// TwinCAT 3 PLC project CartonPLC
// ProgramVersion: 3.1.4026.28
// libraries:
//   SPT Base Types, 3.9.0 (Beckhoff Automation LLC)
//   Tc3_PackML_V2, * (Beckhoff Automation GmbH)
//   Tc3_EventLogger, * (Beckhoff Automation GmbH)
//   Tc2_System, * (Beckhoff Automation GmbH)
//   Tc3_Module, * (Beckhoff Automation GmbH)
//   Tc2_Standard, * (Beckhoff Automation GmbH)
// project tree:
//   / E_ConsoleCommand.TcDUT, GVL_HMI.TcGVL, FB_VirtualCylinder.TcPOU, FB_StrokeStation.TcPOU, FB_CartonCell.TcPOU, FB_SimAxis.TcPOU, FB_SealInspection.TcPOU, FB_CellDevices.TcPOU, I_LineClamp.TcIO, FB_LineClamp.TcPOU, FB_ContinuousLine.TcPOU, FB_LineEvents.TcPOU, MAIN.TcPOU, PlcTask.TcTTO
// real-time tasks:
//   TASK PlcTask: cycle T#10ms, priority 20, ADS port 350

CONFIGURATION CartonPLC
    RESOURCE PLC ON TwinCAT3
        TASK PlcTask(INTERVAL := T#10ms, PRIORITY := 20);
        PROGRAM MAIN WITH PlcTask : MAIN;
    END_RESOURCE
END_CONFIGURATION

// ---- E_ConsoleCommand.TcDUT
{attribute 'qualified_only'}
TYPE E_ConsoleCommand :
(
    Reset := 1,
    Start := 2,
    Hold := 3,
    Unhold := 4,
    Suspend := 5,
    Unsuspend := 6,
    Stop := 7,
    Abort := 8,
    Clear := 9,
    Automatic := 10,
    Manual := 11,
    Stroke1 := 12,
    Stroke2 := 13,
    Stroke3 := 14,
    Stroke4 := 15,
    Stroke5 := 16,
    DropAir := 17,
    RestoreAir := 18,
    LowBlanks := 19,
    Refill := 20,
    MissingSeal := 21,
    RestoreSeal := 22,
    LoopLine := 23,
    Bench := 24,
    Standard := 25,
    Precision := 26,
    JamClamp := 27,
    ReleaseClamp := 28,
    AckClamp := 29
) DINT;
END_TYPE

// ---- GVL_HMI.TcGVL
{attribute 'qualified_only'}
VAR_GLOBAL
    // One atomic DINT per request. See docs/ads.md for the word layout.
    Request : DINT;
    Status : ARRAY[0..105] OF DINT;
END_VAR

// ---- I_LineClamp.TcIO
INTERFACE I_LineClamp

METHOD Follow : DINT
VAR_INPUT
    Extend : BOOL;
END_VAR
END_METHOD

METHOD Home
END_METHOD

END_INTERFACE

// ---- MAIN.TcPOU
PROGRAM MAIN
VAR
    Cell : FB_CartonCell := (Name := 'Carton Cell');
END_VAR

Cell.RunScan();

END_PROGRAM

// ---- FB_CartonCell.TcPOU
FUNCTION_BLOCK FB_CartonCell EXTENDS SPT_BaseTypes.FB_PackML_BaseModule
VAR
    Line : FB_ContinuousLine;
    LineEvents : FB_LineEvents;
    Devices : FB_CellDevices;
    Stations : ARRAY[1..5] OF FB_StrokeStation;
    ActiveStation : DINT;
    Finished : BOOL;
    Cartons : DINT;
    AirFault : BOOL;
    LowStock : BOOL;
    PreviousState : Tc3_PackML_V2.E_PMLState;
    ActingScans : INT;
    RequestSample : DINT;
    Acknowledged : DINT;
    Accepted : BOOL;
    StatusBuffer : ARRAY[0..105] OF DINT;
END_VAR

METHOD PROTECTED Initialize : BOOL
// User mode 4 keeps Idle and Complete for one-station commissioning.
CustomModes(eMode := 4, sName := 'Manual stroke', bDisableHeld := TRUE,
    bDisableSuspended := TRUE, bEnableUnitModeChangeStopped := TRUE);
Initialize := SUPER^.Initialize();
END_METHOD

METHOD RunScan
IF _InitComplete THEN
    CyclicLogic();
ELSE
    _InitComplete := Initialize();
END_IF
END_METHOD

METHOD CyclicLogic
// SPT can call this hook while Initialize is still on the stack.
IF NOT _InitComplete THEN RETURN; END_IF

IF _CurrentState <> PreviousState THEN
    ActingScans := 0;
    PreviousState := _CurrentState;
ELSE
    ActingScans := MIN(45, ActingScans + 1);
END_IF

// Sample once so a concurrent ADS write belongs entirely to one scan.
RequestSample := GVL_HMI.Request;
IF RequestSample <> Acknowledged THEN
    Accepted := ApplyCommand(RequestSample MOD 256);
    Acknowledged := RequestSample;
END_IF

Line.Clock((_CurrentState = Tc3_PackML_V2.E_PMLState.ePMLState_Execute) AND Line.Enabled AND (_CurrentMode = E_PMLUnitMode.ePMLUnitMode_Production));
SUPER^.CyclicLogic();
LineEvents(Occurrence := Line.Occurrence, Alarm := Line.Alarm, Jammed := Line.Jammed,
    Idle := _CurrentState = Tc3_PackML_V2.E_PMLState.ePMLState_Idle);
PublishStatus();
END_METHOD

METHOD PROTECTED Execute
IF Line.Enabled AND (_CurrentMode = E_PMLUnitMode.ePMLUnitMode_Production) THEN
    IF Line.Alarm = 0 THEN Line.Step(Devices.MissingSeal); END_IF
    IF Line.Alarm <> 0 THEN ChangeState(Tc3_PackML_V2.E_PMLCommand.ePMLCommand_Abort); END_IF
    RETURN;
END_IF
IF (ActiveStation < 1) OR (ActiveStation > 5) THEN RETURN; END_IF
IF Finished THEN
    StateComplete();
    RETURN;
END_IF

Stations[ActiveStation].Step();
IF _CurrentMode = E_PMLUnitMode.ePMLUnitMode_Production THEN
    Devices.ProcessStation(ActiveStation, Stations[ActiveStation].Phase);
END_IF

IF Stations[ActiveStation].Done AND
   ((_CurrentMode = E_PMLUnitMode.ePMLUnitMode_UserMode1) OR Devices.ReadyToLeave(ActiveStation)) THEN
    IF (_CurrentMode = E_PMLUnitMode.ePMLUnitMode_UserMode1) OR (ActiveStation = 5) THEN
        Finished := TRUE;
        IF _CurrentMode = E_PMLUnitMode.ePMLUnitMode_Production THEN
            IF Devices.FinishCarton() THEN
                Cartons := Cartons + 1;
            END_IF
        END_IF
        StateComplete();
    ELSIF Devices.IndexToNext(ActiveStation) THEN
        ActiveStation := ActiveStation + 1;
    END_IF
END_IF
END_METHOD

METHOD PROTECTED Resetting
VAR
    StationIndex : INT;
END_VAR
FOR StationIndex := 1 TO 5 DO
    Stations[StationIndex].ResetStation();
END_FOR
Devices.ResetDevices();
Line.ResetLine();
ActiveStation := 0;
Finished := FALSE;
IF (_CurrentState = PreviousState) AND (ActingScans >= 45) THEN
    StateComplete();
END_IF
END_METHOD

METHOD PROTECTED Clearing
IF (_CurrentState = PreviousState) AND (ActingScans >= 45) THEN
    StateComplete();
END_IF
END_METHOD

METHOD PROTECTED Starting
IF (_CurrentState = PreviousState) AND (ActingScans >= 45) THEN
    StateComplete();
END_IF
END_METHOD

METHOD PROTECTED Stopping
IF (_CurrentState = PreviousState) AND (ActingScans >= 45) THEN
    StateComplete();
END_IF
END_METHOD

METHOD PROTECTED Aborting
IF (_CurrentState = PreviousState) AND (ActingScans >= 45) THEN
    StateComplete();
END_IF
END_METHOD

METHOD PROTECTED Holding
IF (_CurrentState = PreviousState) AND (ActingScans >= 45) THEN
    StateComplete();
END_IF
END_METHOD

METHOD PROTECTED Unholding
IF (_CurrentState = PreviousState) AND (ActingScans >= 45) THEN
    StateComplete();
END_IF
END_METHOD

METHOD PROTECTED Suspending
IF (_CurrentState = PreviousState) AND (ActingScans >= 45) THEN
    StateComplete();
END_IF
END_METHOD

METHOD PROTECTED Unsuspending
IF (_CurrentState = PreviousState) AND (ActingScans >= 45) THEN
    StateComplete();
END_IF
END_METHOD

METHOD PROTECTED Completing
IF (_CurrentState = PreviousState) AND (ActingScans >= 45) THEN
    StateComplete();
END_IF
END_METHOD

METHOD PRIVATE ApplyCommand : BOOL
VAR_INPUT
    Code : DINT;
END_VAR
VAR
    IsManual : BOOL;
END_VAR
IsManual := _CurrentMode = E_PMLUnitMode.ePMLUnitMode_UserMode1;
CASE Code OF
    E_ConsoleCommand.Reset:
        IF NOT AirFault AND ((_CurrentState = Tc3_PackML_V2.E_PMLState.ePMLState_Stopped) OR (_CurrentState = Tc3_PackML_V2.E_PMLState.ePMLState_Complete)) THEN
            ChangeState(Tc3_PackML_V2.E_PMLCommand.ePMLCommand_Reset);
            ApplyCommand := TRUE;
        END_IF
    E_ConsoleCommand.Start:
        IF NOT IsManual AND (_CurrentState = Tc3_PackML_V2.E_PMLState.ePMLState_Idle) THEN
            Line.Timing := Line.Enabled;
            ActiveStation := SEL(Line.Enabled, 1, 0);
            ChangeState(Tc3_PackML_V2.E_PMLCommand.ePMLCommand_Start);
            ApplyCommand := TRUE;
        END_IF
    E_ConsoleCommand.Hold:
        IF NOT IsManual AND (_CurrentState = Tc3_PackML_V2.E_PMLState.ePMLState_Execute) THEN
            ChangeState(Tc3_PackML_V2.E_PMLCommand.ePMLCommand_Hold);
            ApplyCommand := TRUE;
        END_IF
    E_ConsoleCommand.Unhold:
        IF _CurrentState = Tc3_PackML_V2.E_PMLState.ePMLState_Held THEN
            ChangeState(Tc3_PackML_V2.E_PMLCommand.ePMLCommand_Unhold);
            ApplyCommand := TRUE;
        END_IF
    E_ConsoleCommand.Suspend:
        IF NOT IsManual AND (_CurrentState = Tc3_PackML_V2.E_PMLState.ePMLState_Execute) THEN
            ChangeState(Tc3_PackML_V2.E_PMLCommand.ePMLCommand_Suspend);
            ApplyCommand := TRUE;
        END_IF
    E_ConsoleCommand.Unsuspend:
        IF _CurrentState = Tc3_PackML_V2.E_PMLState.ePMLState_Suspended THEN
            ChangeState(Tc3_PackML_V2.E_PMLCommand.ePMLCommand_Unsuspend);
            ApplyCommand := TRUE;
        END_IF
    E_ConsoleCommand.Stop:
        IF (_CurrentState <> Tc3_PackML_V2.E_PMLState.ePMLState_Undefined) AND
            (_CurrentState <> Tc3_PackML_V2.E_PMLState.ePMLState_Stopped) AND
            (_CurrentState <> Tc3_PackML_V2.E_PMLState.ePMLState_Stopping) AND
            (_CurrentState <> Tc3_PackML_V2.E_PMLState.ePMLState_Aborted) AND
            (_CurrentState <> Tc3_PackML_V2.E_PMLState.ePMLState_Aborting) AND
            (_CurrentState <> Tc3_PackML_V2.E_PMLState.ePMLState_Clearing) THEN
            Line.Timing := FALSE;
            ChangeState(Tc3_PackML_V2.E_PMLCommand.ePMLCommand_Stop);
            ApplyCommand := TRUE;
        END_IF
    E_ConsoleCommand.Abort:
        IF (_CurrentState <> Tc3_PackML_V2.E_PMLState.ePMLState_Aborted) AND
            (_CurrentState <> Tc3_PackML_V2.E_PMLState.ePMLState_Aborting) AND
            (_CurrentState <> Tc3_PackML_V2.E_PMLState.ePMLState_Undefined) THEN
            ChangeState(Tc3_PackML_V2.E_PMLCommand.ePMLCommand_Abort);
            ApplyCommand := TRUE;
        END_IF
    E_ConsoleCommand.Clear:
        IF NOT AirFault AND ((Line.Alarm = 0) OR ((Line.Alarm = 2) AND NOT Line.Jammed)) AND (_CurrentState = Tc3_PackML_V2.E_PMLState.ePMLState_Aborted) THEN
            Line.ClearAlarm();
            ChangeState(Tc3_PackML_V2.E_PMLCommand.ePMLCommand_Clear);
            ApplyCommand := TRUE;
        END_IF
    E_ConsoleCommand.Manual, E_ConsoleCommand.Automatic:
        IF _CurrentState = Tc3_PackML_V2.E_PMLState.ePMLState_Stopped THEN
            IF (Code = E_ConsoleCommand.Manual) AND NOT IsManual THEN
                Line.Timing := FALSE;
                ChangeMode(E_PMLUnitMode.ePMLUnitMode_UserMode1);
                ApplyCommand := TRUE;
            ELSIF (Code = E_ConsoleCommand.Automatic) AND IsManual THEN
                ChangeMode(E_PMLUnitMode.ePMLUnitMode_Production);
                ApplyCommand := TRUE;
            END_IF
        END_IF
    E_ConsoleCommand.Stroke1..E_ConsoleCommand.Stroke5:
        IF IsManual AND (_CurrentState = Tc3_PackML_V2.E_PMLState.ePMLState_Idle) THEN
            ActiveStation := Code - E_ConsoleCommand.Stroke1 + 1;
            ChangeState(Tc3_PackML_V2.E_PMLCommand.ePMLCommand_Start);
            ApplyCommand := TRUE;
        END_IF
    E_ConsoleCommand.DropAir:
        ApplyCommand := NOT AirFault;
        AirFault := TRUE;
        IF (_CurrentState <> Tc3_PackML_V2.E_PMLState.ePMLState_Aborted) AND (_CurrentState <> Tc3_PackML_V2.E_PMLState.ePMLState_Aborting) THEN
            ChangeState(Tc3_PackML_V2.E_PMLCommand.ePMLCommand_Abort);
        END_IF
    E_ConsoleCommand.RestoreAir:
        ApplyCommand := AirFault;
        AirFault := FALSE;
    E_ConsoleCommand.LowBlanks:
        ApplyCommand := NOT LowStock;
        LowStock := TRUE;
    E_ConsoleCommand.MissingSeal:
        ApplyCommand := NOT Devices.MissingSeal;
        Devices.MissingSeal := TRUE;
    E_ConsoleCommand.RestoreSeal:
        ApplyCommand := Devices.MissingSeal;
        Devices.MissingSeal := FALSE;
    E_ConsoleCommand.LoopLine, E_ConsoleCommand.Bench:
        IF NOT IsManual AND (_CurrentState = Tc3_PackML_V2.E_PMLState.ePMLState_Stopped) THEN
            ApplyCommand := Line.Enabled <> (Code = E_ConsoleCommand.LoopLine);
            Line.Timing := FALSE;
            Line.Enabled := Code = E_ConsoleCommand.LoopLine;
        END_IF
    E_ConsoleCommand.Standard, E_ConsoleCommand.Precision:
        IF Line.Enabled AND NOT IsManual AND (_CurrentState = Tc3_PackML_V2.E_PMLState.ePMLState_Stopped) THEN
            ApplyCommand := Line.Precision <> (Code = E_ConsoleCommand.Precision);
            Line.Precision := Code = E_ConsoleCommand.Precision;
        END_IF
    E_ConsoleCommand.JamClamp:
        IF Line.Enabled AND NOT IsManual AND NOT Line.Jammed AND (Line.Alarm = 0) THEN
            Line.Jammed := TRUE; ApplyCommand := TRUE;
        END_IF
    E_ConsoleCommand.ReleaseClamp:
        ApplyCommand := Line.Jammed; Line.Jammed := FALSE;
    E_ConsoleCommand.AckClamp:
        IF (_CurrentState = Tc3_PackML_V2.E_PMLState.ePMLState_Aborted) AND
            (Line.Alarm = 1) AND (RequestSample / 256 = Line.Occurrence) THEN
            Line.AcknowledgeAlarm(); ApplyCommand := TRUE;
        END_IF
    E_ConsoleCommand.Refill:
        ApplyCommand := LowStock;
        LowStock := FALSE;
END_CASE
END_METHOD

METHOD PRIVATE PublishStatus
StatusBuffer[0] := 51003;
StatusBuffer[1] := TO_DINT(_CurrentState);
StatusBuffer[2] := BOOL_TO_DINT(_CurrentMode = E_PMLUnitMode.ePMLUnitMode_UserMode1);
StatusBuffer[3] := ActiveStation;
StatusBuffer[4] := 0;
IF (ActiveStation >= 1) AND (ActiveStation <= 5) THEN
    StatusBuffer[4] := Stations[ActiveStation].Phase;
END_IF
StatusBuffer[5] := Cartons;
StatusBuffer[6] := BOOL_TO_DINT(AirFault);
StatusBuffer[7] := BOOL_TO_DINT(LowStock);
StatusBuffer[8] := Acknowledged;
StatusBuffer[9] := (StatusBuffer[9] MOD 2000000000) + 1;
StatusBuffer[10] := BOOL_TO_DINT(Accepted);
Devices.Publish(StatusBuffer);
Line.Publish(StatusBuffer);
GVL_HMI.Status := StatusBuffer;
END_METHOD

END_FUNCTION_BLOCK

// ---- FB_ContinuousLine.TcPOU
FUNCTION_BLOCK FB_ContinuousLine
VAR
    Clamp : FB_LineClamp;
    Actuator : I_LineClamp;
    Vision : FB_SealInspection;
    Products, Checks, Failures : ARRAY[0..15] OF DINT;
    CamX, CamZ : ARRAY[0..7] OF DINT;
    Tick, PitchIndex, Issued, Good, Rejected, LastId, LastFailed, LastChecked, Discarded : DINT;
    RunTicks, PlannedTicks, IdealTicks, WaitTicks, Travel, ClampMm : DINT;
    ClampRequest : BOOL;
END_VAR
VAR_INPUT
    Enabled : BOOL := TRUE;
    Precision, Jammed, Timing : BOOL;
END_VAR
VAR_OUTPUT
    Alarm, Occurrence : DINT;
END_VAR

METHOD ClearAlarm
Alarm := 0;
END_METHOD

METHOD AcknowledgeAlarm
Alarm := 2;
END_METHOD

METHOD Clock
VAR_INPUT
    Executing : BOOL;
END_VAR
IF Timing THEN
    PlannedTicks := PlannedTicks + 1;
    IF Executing THEN RunTicks := RunTicks + 1; END_IF
END_IF
END_METHOD

METHOD ResetLine
VAR
    i : INT;
END_VAR
FOR i := 0 TO 15 DO
    IF Products[i] <> 0 THEN Discarded := Discarded + 1; END_IF
    Products[i] := 0; Checks[i] := 0; Failures[i] := 0;
END_FOR
FOR i := 0 TO 7 DO CamX[i] := 0; CamZ[i] := 0; END_FOR
Tick := 0; PitchIndex := 0; WaitTicks := 0; Travel := 0;
Actuator := Clamp;
Actuator.Home();
ClampMm := 0; ClampRequest := FALSE;
END_METHOD

METHOD AtSlot : DINT
VAR_INPUT
    Slot, Count : DINT;
END_VAR
AtSlot := (Slot + Count - (PitchIndex MOD Count)) MOD Count;
END_METHOD

METHOD Ease : DINT
VAR_INPUT
    InputPhase : DINT;
END_VAR
VAR
    u : DINT;
END_VAR
u := LIMIT(0, InputPhase, 100);
Ease := u * u * (300 - 2 * u) / 1000;
END_METHOD

METHOD InspectMover
VAR_INPUT
    Mover, BitNumber : DINT;
    Passed : BOOL;
END_VAR
VAR
    Mask : DWORD;
END_VAR
Mask := SHL(DWORD#1, DINT_TO_UINT(BitNumber));
Checks[Mover] := DWORD_TO_DINT(DINT_TO_DWORD(Checks[Mover]) OR Mask);
IF NOT Passed THEN Failures[Mover] := DWORD_TO_DINT(DINT_TO_DWORD(Failures[Mover]) OR Mask); END_IF
END_METHOD

METHOD Step
VAR_INPUT
    MissingSeal : BOOL;
END_VAR
VAR
    p, Mover, Station, Reach, Depth, Stroke : DINT;
    FirstScan : BOOL;
END_VAR
VAR CONSTANT
    Period : DINT := 200; // 2 s at the 10 ms scan rate
END_VAR
Stroke := SEL(Precision, 40, 48);
p := Tick * 100 / Period;
FirstScan := (Tick MOD (Period / 100)) = 0;
Mover := AtSlot(0, 10);
IF (Tick = 0) AND (Products[Mover] = 0) THEN
    Issued := Issued + 1; Products[Mover] := Issued;
END_IF
ClampRequest := (Products[AtSlot(2, 10)] <> 0) AND (p >= 12) AND (p < 54);
Actuator := Clamp;
Clamp.Jammed := Jammed;
ClampMm := Actuator.Follow(ClampRequest);
IF ClampRequest AND (ClampMm < 16) THEN WaitTicks := WaitTicks + 1; ELSE WaitTicks := 0; END_IF
IF WaitTicks >= 15 THEN
    Occurrence := (Occurrence MOD 8388606) + 1;
    Alarm := 1;
    RETURN;
END_IF
IF p < 12 THEN Reach := Ease(p * 100 / 12);
ELSIF p < 48 THEN Reach := 1000;
ELSE Reach := 1000 - Ease((p - 48) * 100 / 12); END_IF
IF p < 12 THEN Depth := 0;
ELSIF p < 26 THEN Depth := Ease((p - 12) * 100 / 14);
ELSIF p < 36 THEN Depth := 1000;
ELSE Depth := 1000 - Ease((p - 36) * 100 / 12); END_IF
Travel := Ease((p - 60) * 100 / 40);
FOR Station := 0 TO 7 DO
    Mover := AtSlot(SEL(Station < 4, Station + 1, Station), 10);
    IF Products[Mover] <> 0 THEN
        CamX[Station] := Reach * (100 + Station * 4) / 1000;
        CamZ[Station] := Depth * Stroke / 1000;
        IF Station = 5 THEN
            IF p <= 80 THEN CamX[Station] := Travel / 2;
            ELSE CamX[Station] := 250 - Ease((p-80)*100/20) / 4; END_IF
            IF p < 60 THEN CamZ[Station] := 0;
            ELSIF p <= 74 THEN CamZ[Station] := Ease((p-60)*100/14) * Stroke / 1000;
            ELSE CamZ[Station] := (1000-Ease((p-78)*100/8)) * Stroke / 1000; END_IF
        END_IF
        IF (p = SEL(Station = 5, 32, 76)) AND FirstScan THEN
            InspectMover(Mover, Station, (CamZ[Station] = Stroke) AND ((Station <> 2) OR (ClampMm = 16)));
        END_IF
    ELSE CamX[Station] := 0; CamZ[Station] := 0; END_IF
END_FOR
IF (p = 54) AND FirstScan THEN ProcessTable(MissingSeal, Period); END_IF
Tick := Tick + 1;
IF Tick = Period THEN
    Tick := 0; Travel := 0; PitchIndex := (PitchIndex + 1) MOD 30;
END_IF
END_METHOD

METHOD ProcessTable
VAR_INPUT
    MissingSeal : BOOL;
    Period : DINT;
END_VAR
VAR
    Source, Target, Seat, Camera, Pack : DINT;
END_VAR
Source := AtSlot(8,10); Target := 10 + AtSlot(0,6);
IF (Products[Source] <> 0) AND (Products[Target] = 0) THEN
    Products[Target] := Products[Source]; Checks[Target] := Checks[Source]; Failures[Target] := Failures[Source];
    Products[Source] := 0; Checks[Source] := 0; Failures[Source] := 0;
END_IF
Seat := 10 + AtSlot(1,6); Camera := 10 + AtSlot(2,6); Pack := 10 + AtSlot(3,6);
IF Products[Seat] <> 0 THEN InspectMover(Seat, 8, (DINT_TO_DWORD(Checks[Seat]) AND DWORD#255) = DWORD#255); END_IF
IF Products[Camera] <> 0 THEN
    Vision.ClearResult(); Vision.Inspect(MissingSeal);
    InspectMover(Camera, 9, Vision.Verdict = 1);
END_IF
IF Products[Pack] <> 0 THEN
    LastId := Products[Pack]; LastChecked := Checks[Pack]; LastFailed := Failures[Pack];
    IF (LastChecked = 1023) AND (LastFailed = 0) THEN Good := Good + 1;
    ELSE Rejected := Rejected + 1; END_IF
    IdealTicks := IdealTicks + Period;
    Products[Pack] := 0; Checks[Pack] := 0; Failures[Pack] := 0;
END_IF
END_METHOD

METHOD Publish
VAR_IN_OUT
    Words : ARRAY[0..105] OF DINT;
END_VAR
VAR
    i : INT;
END_VAR
Words[20] := BOOL_TO_DINT(Enabled);
Words[21] := BOOL_TO_DINT(Precision);
Words[22] := Tick;
Words[23] := PitchIndex;
Words[24] := Issued;
Words[25] := Good;
Words[26] := Rejected;
Words[27] := LastId;
Words[28] := LastFailed;
Words[29] := BOOL_TO_DINT(Jammed);
Words[30] := Occurrence;
Words[31] := Alarm;
Words[32] := BOOL_TO_DINT(ClampRequest);
Words[33] := ClampMm;
Words[34] := RunTicks;
Words[35] := PlannedTicks;
Words[36] := IdealTicks;
Words[37] := Discarded;
FOR i := 0 TO 15 DO
    Words[40+i] := Products[i]; Words[56+i] := Checks[i]; Words[72+i] := Failures[i];
END_FOR
FOR i := 0 TO 7 DO Words[88+i] := CamX[i]; Words[96+i] := CamZ[i]; END_FOR
Words[104] := Travel;
Words[105] := LastChecked;
END_METHOD

END_FUNCTION_BLOCK

// ---- FB_LineClamp.TcPOU
FUNCTION_BLOCK FB_LineClamp IMPLEMENTS I_LineClamp
VAR_INPUT
    Jammed : BOOL;
END_VAR
VAR
    Position : DINT;
END_VAR

METHOD Follow : DINT
VAR_INPUT
    Extend : BOOL;
END_VAR
IF NOT Extend THEN Position := MAX(0, Position - 4);
ELSIF NOT Jammed THEN Position := MIN(16, Position + 4);
END_IF
Follow := Position;
END_METHOD

METHOD Home
Position := 0;
END_METHOD

END_FUNCTION_BLOCK

// ---- FB_SealInspection.TcPOU
FUNCTION_BLOCK FB_SealInspection
VAR_OUTPUT
    Verdict : DINT; // 0 pending, 1 pass, 2 reject
    BrightSamples : DINT;
END_VAR
VAR CONSTANT
    GoodPixels : ARRAY[0..4] OF USINT := [231, 236, 228, 239, 232];
    MissingPixels : ARRAY[0..4] OF USINT := [118, 122, 120, 124, 121];
END_VAR

METHOD Inspect
VAR_INPUT
    MissingSeal : BOOL;
END_VAR
VAR
    Index : INT;
    Pixel : USINT;
END_VAR
IF Verdict <> 0 THEN RETURN; END_IF
FOR Index := 0 TO 4 DO
    Pixel := SEL(MissingSeal, GoodPixels[Index], MissingPixels[Index]);
    IF Pixel >= 200 THEN
        BrightSamples := BrightSamples + 1;
    END_IF
END_FOR
Verdict := SEL(BrightSamples >= 4, 2, 1);
END_METHOD

METHOD ClearResult
Verdict := 0;
BrightSamples := 0;
END_METHOD

END_FUNCTION_BLOCK

// ---- FB_LineEvents.TcPOU
FUNCTION_BLOCK FB_LineEvents
VAR_INPUT
    Occurrence, Alarm : DINT;
    Jammed, Idle : BOOL;
END_VAR
VAR
    Event : Tc3_EventLogger.FB_TcAlarm;
    Recovery : Tc3_EventLogger.FB_TcMessage;
    Created, MessageCreated, Confirmed, Cleared, Recovered : BOOL;
    Seen : DINT;
END_VAR

IF NOT Created THEN Created := Event.CreateEx(TC_EVENTS.CartonLine.ClampTimeout, TRUE, 0) = 0; END_IF
IF NOT MessageCreated THEN MessageCreated := Recovery.CreateEx(TC_EVENTS.CartonLine.LineRecovered, 0) = 0; END_IF
IF Created AND (Occurrence <> Seen) THEN
    Event.ipArguments.Clear().AddDInt(Occurrence);
    IF Event.Raise(0) = 0 THEN Seen := Occurrence; Confirmed := FALSE; Cleared := FALSE; Recovered := FALSE; END_IF
END_IF
IF (Seen <> 0) AND (Seen = Occurrence) THEN
    IF (Alarm = 2) AND NOT Confirmed THEN Confirmed := Event.Confirm(0) = 0; END_IF
    IF NOT Jammed AND NOT Cleared THEN Cleared := Event.Clear(0, FALSE) = 0; END_IF
    IF MessageCreated AND Idle AND (Alarm = 0) AND NOT Recovered THEN
        Recovery.ipArguments.Clear().AddDInt(Occurrence);
        Recovered := Recovery.Send(0) = 0;
    END_IF
END_IF

END_FUNCTION_BLOCK

// ---- FB_CellDevices.TcPOU
FUNCTION_BLOCK FB_CellDevices
VAR
    FeedAxis : FB_SimAxis;
    TrackMover : FB_SimAxis;
    ShuttleX : FB_SimAxis;
    ShuttleY : FB_SimAxis;
    Camera : FB_SealInspection;
END_VAR
VAR_OUTPUT
    Indexing : BOOL;
    Rejected : DINT;
END_VAR
VAR_INPUT
    MissingSeal : BOOL;
END_VAR

METHOD ResetDevices
FeedAxis.Home();
TrackMover.Home();
ShuttleX.Home();
ShuttleY.Home();
Camera.ClearResult();
Indexing := FALSE;
END_METHOD

METHOD ProcessStation
VAR_INPUT
    Station : DINT;
    Phase : DINT;
END_VAR
CASE Station OF
    1: // Servo meters a 180 mm blank.
        FeedAxis.MoveToward(180, 2);
    4: // Trigger once when the closing platen reaches its forward limit.
        IF Phase >= 100 THEN Camera.Inspect(MissingSeal); END_IF
    5: // Route the sealed carton to one of two discharge lanes.
        ShuttleX.MoveToward(240, 2);
        ShuttleY.MoveToward(SEL(Camera.Verdict = 1, -120, 120), 2);
END_CASE
END_METHOD

METHOD IndexToNext : BOOL
VAR_INPUT
    Station : DINT;
END_VAR
IndexToNext := TrackMover.MoveToward(Station * 560, 8);
Indexing := NOT IndexToNext;
END_METHOD

METHOD ReadyToLeave : BOOL
VAR_INPUT
    Station : DINT;
END_VAR
CASE Station OF
    1: ReadyToLeave := FeedAxis.PositionMm = 180;
    4: ReadyToLeave := Camera.Verdict <> 0;
    5: ReadyToLeave := (ShuttleX.PositionMm = 240) AND
           (ShuttleY.PositionMm = SEL(Camera.Verdict = 1, -120, 120));
ELSE
    ReadyToLeave := TRUE;
END_CASE
END_METHOD

METHOD FinishCarton : BOOL
FinishCarton := Camera.Verdict = 1;
IF NOT FinishCarton THEN Rejected := Rejected + 1; END_IF
END_METHOD

METHOD Publish
VAR_IN_OUT
    Words : ARRAY[0..105] OF DINT;
END_VAR
Words[11] := FeedAxis.PositionMm;
Words[12] := TrackMover.PositionMm;
Words[13] := ShuttleX.PositionMm;
Words[14] := ShuttleY.PositionMm;
Words[15] := Camera.Verdict;
Words[16] := Rejected;
Words[17] := BOOL_TO_DINT(MissingSeal);
Words[18] := BOOL_TO_DINT(Indexing);
Words[19] := Camera.BrightSamples;
END_METHOD

END_FUNCTION_BLOCK

// ---- FB_SimAxis.TcPOU
FUNCTION_BLOCK FB_SimAxis
VAR_OUTPUT
    PositionMm : DINT;
END_VAR

METHOD MoveToward : BOOL
VAR_INPUT
    TargetMm : DINT;
    MaxStepMm : DINT;
END_VAR
// Deterministic virtual axis. One invocation corresponds to one 10 ms task tick.
PositionMm := PositionMm + LIMIT(-MaxStepMm, TargetMm - PositionMm, MaxStepMm);
MoveToward := PositionMm = TargetMm;
END_METHOD

METHOD Home
PositionMm := 0;
END_METHOD

END_FUNCTION_BLOCK

// ---- FB_StrokeStation.TcPOU
FUNCTION_BLOCK FB_StrokeStation
VAR_OUTPUT
    Phase : DINT; // Outstroke 0..100, return 101..200
    Done : BOOL;
END_VAR
VAR
    Cylinder : FB_VirtualCylinder;
    Returning : BOOL;
END_VAR

METHOD ResetStation
Cylinder.Home();
Returning := FALSE;
Phase := 0;
Done := FALSE;
END_METHOD

METHOD Step
IF Done THEN RETURN; END_IF
Cylinder.FollowStroke(Forward := NOT Returning);
IF Returning THEN
    Phase := 200 - Cylinder.Position;
    Done := Cylinder.Position = 0;
ELSE
    Phase := Cylinder.Position;
    Returning := Cylinder.Position = 100;
END_IF
END_METHOD

END_FUNCTION_BLOCK

// ---- FB_VirtualCylinder.TcPOU
FUNCTION_BLOCK FB_VirtualCylinder
VAR_OUTPUT
    Position : DINT; // 0 = home, 100 = forward limit
END_VAR

METHOD FollowStroke
VAR_INPUT
    Forward : BOOL;
END_VAR
IF Forward THEN
    Position := MIN(100, Position + 1);
ELSE
    Position := MAX(0, Position - 1);
END_IF
END_METHOD

METHOD Home
Position := 0;
END_METHOD

END_FUNCTION_BLOCK
